FUNCTION_BLOCK InOut4
  (* Standard: 61499-1; Description: Copyright (c) 2026 Martin Erich Jobst This program and the accompanying materials are made available under the terms of the Eclipse Public License 2.0 which is available at https://www.eclipse.org/legal/epl-2.0/ SPDX-License-Identifier: EPL-2.0 *)
  (* Version 1.0, 2026-11-18, Martin Jobst *)
  PACKAGE lib::VarDeclaration::support;
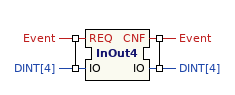
  EVENT_INPUT
    REQ WITH IO;
  END_EVENT
  EVENT_OUTPUT
    CNF WITH IO;
  END_EVENT
  VAR_IN_OUT
    IO : ARRAY [0..3] OF DINT;
  END_VAR
END_FUNCTION_BLOCK
